DATA_BLOCK "GDB_FrameProbe"
{ S7_Optimized_Access := 'TRUE' }
VERSION : 0.1
NON_RETAIN
VAR
    Order : DInt;
    Scans : DInt;
    Checks : DInt;
    FailedChecks : DInt;
    Passed : Bool;
    OverflowPassed : Bool;
    BadParentPassed : Bool;
    Rows : Array[0..16] of "FRK_ProbeRow";
END_VAR
BEGIN
END_DATA_BLOCK
